FUNCTION_BLOCK FB_SwitchMonostable IMPLEMENTS I_Switch
VAR_INPUT
    stDeviceId : ST_DeviceId;
    bInput     : BOOL;
END_VAR
VAR
    bPreviousInput : BOOL;
    bPressed       : BOOL;
    bReleased      : BOOL;
END_VAR

bPressed := bInput AND NOT bPreviousInput;
bReleased := NOT bInput AND bPreviousInput;

bPreviousInput := bInput;

PROPERTY DeviceId : ST_DeviceId
GET
DeviceId := stDeviceId;
END_GET
END_PROPERTY

PROPERTY IsPressed : BOOL
GET
IsPressed := bInput;
END_GET
END_PROPERTY

PROPERTY Pressed : BOOL
GET
Pressed := bPressed;
END_GET
END_PROPERTY

PROPERTY Released : BOOL
GET
Released := bReleased;
END_GET
END_PROPERTY

END_FUNCTION_BLOCK

(* stored: Version 1.1.0.1, ProductVersion 3.1.4026.20
   POU FB_SwitchMonostable: Id {7B1F2D31-7A6B-4C2D-9F31-2A8C5D1E2001}
   Property DeviceId: Id {7B1F2D31-7A6B-4C2D-9F31-2A8C5D1E2011}
   Get Get: Id {7B1F2D31-7A6B-4C2D-9F31-2A8C5D1E2012}
   Property IsPressed: Id {7B1F2D31-7A6B-4C2D-9F31-2A8C5D1E2021}
   Get Get: Id {7B1F2D31-7A6B-4C2D-9F31-2A8C5D1E2022}
   Property Pressed: Id {7B1F2D31-7A6B-4C2D-9F31-2A8C5D1E2031}
   Get Get: Id {7B1F2D31-7A6B-4C2D-9F31-2A8C5D1E2032}
   Property Released: Id {7B1F2D31-7A6B-4C2D-9F31-2A8C5D1E2041}
   Get Get: Id {7B1F2D31-7A6B-4C2D-9F31-2A8C5D1E2042} *)
